TYPE ET_GFX4IR_1 :
(
	ET_GFX4IRState_eWaitExecute := 0,
	ET_GFX4IRState_eCtrlOn,
	ET_GFX4IRState_eCtrlOff,
	ET_GFX4IRState_eDone := 197,
	ET_GFX4IRState_eError := 198,
	ET_GFX4IRState_eNoExecute := 199
);
END_TYPE

(* stored: Version 1.1.0.1, ProductVersion 3.1.4024.15
   DUT ET_GFX4IR_1: Id {2ac6cdbd-996e-49ac-9bb0-79ac2246522e} *)
